TYPE ST_TimeHoursCounter :
STRUCT
	lrAllOverHours					:LREAL; 							(* All over counter hours *)
	lrAfterResetHours					:LREAL; 							(* Counter hours since last reset *)
END_STRUCT
END_TYPE

(* stored: Version 1.1.0.1, ProductVersion 3.1.4024.15
   DUT ST_TimeHoursCounter: Id {e78df8fd-9137-45a8-ab9b-2b5f3bbb5927} *)
